(* IEC 61131-3 sources: volt/packages/volt-lsp-iec/test-corpus/bakon-nano/Device/Plc Logic/Application/Library Manager/CAA Callback Extern, 38 files *)

(* ---- CALLBACK.dut ---- *)
TYPE CALLBACK : CB_CALLBACK;
END_TYPE

(* ---- CB_CALLBACK.dut ---- *)
TYPE CB_CALLBACK :
STRUCT
	PPOUFUNC : CAA.PVOID := CAA.gc_pNULL;
	EEVENT : EVENT := EVENT.ALL_EVENTS;
	ECLASS : EVENT_CLASS := EVENT_CLASS.NO_CLASS;
	ESOURCE : EVENT_SOURCE := EVENT_SOURCE.NO_SOURCE;
END_STRUCT
END_TYPE

(* ---- ERROR.dut ---- *)
TYPE ERROR :
(
	NO_ERROR := 0,
	FIRST_ERROR := 20000,
	HANDLE_INVALID := 20001,
	UNKNOWN_EVENT := 20002,
	CALLBACK_NOT_REMOVABLE := 20003,
	WRONG_ARGUMENT := 20004,
	CB_NO_MEMORY := 20005,
	CB_EVENT_EXISTS := 20006,
	CB_CALL_CALLBACKS_FAILED := 20007,
	CB_NO_SYSTEM_EVENT := 20008,
	CB_BUFFER_NOT_AVAILABLE := 20009,
	CB_SYSTEM_EVENT := 20010,
	FIRST_MF := 20050,
	LAST_ERROR := 20099
);
END_TYPE

(* ---- EVENT.dut ---- *)
TYPE EVENT :
(
	ALL_EVENTS := -1,
	NO_EVENT := 0,
	START := 1000,
	STOP,
	BEFORE_RESET,
	AFTER_RESET,
	SHUTDOWN,
	ONLINE_CHANGE,
	BEFORE_DOWNLOAD,
	TASKCODE_NOT_CALLED,
	TIMER,
	DEBUG_LOOP,
	SCHEDULE,
	ERR_WATCHDOG := 4000,
	ERR_HARDWARE_WATCHDOG,
	ERR_FIELDBUS,
	ERR_IOUPDATE,
	ERR_POWERFAIL,
	EXCPT_ILLEGAL_INSTRUCTION := 5000,
	EXCPT_ACCESS_VIOLATION,
	EXCPT_PRIV_INSTRUCTION,
	EXCPT_IN_PAGE_ERROR,
	EXCPT_STACK_OVERFLOW,
	EXCPT_MISALIGNMENT,
	EXCPT_ARRAYBOUNDS,
	EXCPT_DIVIDEBYZERO,
	EXCPT_OVERFLOW,
	EXCPT_NONCONTINUABLE,
	EXCPT_NO_FPU_AVAILABLE := 5500,
	EXCPT_FPU_ERROR,
	EXCPT_FPU_DENORMAL_OPERAND,
	EXCPT_FPU_DIVIDEBYZERO,
	EXCPT_FPU_INVALID_OPERATION,
	EXCPT_FPU_OVERFLOW,
	EXCPT_FPU_STACK_CHECK,
	INTERRUPT_0 := 6000,
	INTERRUPT_1,
	INTERRUPT_2,
	INTERRUPT_3,
	INTERRUPT_4,
	INTERRUPT_5,
	INTERRUPT_6,
	INTERRUPT_7,
	INTERRUPT_8,
	INTERRUPT_9,
	INTERRUPT_10,
	INTERRUPT_11,
	INTERRUPT_12,
	INTERRUPT_13,
	INTERRUPT_14,
	INTERRUPT_15,
	INTERRUPT_255 := 6255,
	AFTER_READING_INPUTS := 7000,
	BEFORE_WRITING_OUTPUTS,
	TIMER_0 := 9900,
	TIMER_1,
	TIMER_2,
	TIMER_3,
	TIMER_4,
	TIMER_5,
	TIMER_6,
	TIMER_7,
	TIMER_8,
	TIMER_9,
	TIMER_10,
	TIMER_11,
	TIMER_12,
	TIMER_13,
	TIMER_14,
	TIMER_15,
	TIMER_99 := 9999
);
END_TYPE

(* ---- EVENT_CLASS.dut ---- *)
TYPE EVENT_CLASS :
(
	ALL_CLASSES := -1,
	NO_CLASS := 16#0,
	ONLINE_EVENTS := 16#1,
	INFOS := 16#2,
	WARNINGS := 16#4,
	RTS_ERRORS := 16#8,
	SYSTEM_EXCEPTIONS := 16#10,
	INTERRUPTS := 16#20,
	IO := 16#40,
	FIELDBUS := 16#80,
	TIMERS := 16#100,
	MANUF_SPEC := 16#200
);
END_TYPE

(* ---- EVENT_SOURCE.dut ---- *)
TYPE EVENT_SOURCE :
(
	ALL_SOURCES := -1,
	NO_SOURCE := 0,
	RUNTIME := 16#1,
	SYSTEM := 16#2,
	IECTASK := 16#4,
	IECPROGRAM := 16#8,
	DRIVER := 16#10
);
END_TYPE

(* ---- GLOBALCONSTANTS.gvl ---- *)
VAR_GLOBAL
	GC_CBNULL : CB_CALLBACK := STRUCT(pPOUFunc := CAA.gc_pNULL, eEvent := EVENT.NO_EVENT, eClass := EVENT_CLASS.NO_CLASS, eSource := EVENT_SOURCE.NO_SOURCE);
END_VAR

(* ---- RSHANDLING.gvl ---- *)
VAR_GLOBAL
	G_CALLBACKCLASS : CallbackClass;
END_VAR

(* ---- VERSIONCONSTANTS.gvl ---- *)
VAR_GLOBAL
	GC_BYVERSION : BYTE := 1;
	GC_VERSION_1 : BYTE := 0;
END_VAR

(* ---- _CALLFUNCTIONBYINDEX.pou ---- *)
FUNCTION _CALLFUNCTIONBYINDEX : __XWORD
VAR_INPUT
	PPOUFUNC : CAA.PVOID;
	DWPARAM1 : __XWORD;
	DWPARAM2 : __XWORD;
	DWPARAM3 : __XWORD;
	PEERROR : POINTER TO ERROR;
END_VAR
END_FUNCTION

(* ---- _DECODECLASS.pou ---- *)
FUNCTION _DECODECLASS : EVENT_CLASS
VAR_INPUT
	DWSPEC : DWORD;
END_VAR
END_FUNCTION

(* ---- _DECODEEVENT.pou ---- *)
FUNCTION _DECODEEVENT : EVENT
VAR_INPUT
	DWSPEC : DWORD;
END_VAR
END_FUNCTION

(* ---- _ENCODESPEC.pou ---- *)
FUNCTION _ENCODESPEC : DWORD
VAR_INPUT
	EEVENT : EVENT;
	ECLASS : EVENT_CLASS;
END_VAR
END_FUNCTION

(* ---- _GETCALLBACK.pou ---- *)
FUNCTION _GETCALLBACK : ERROR
VAR_INPUT
	HHANDLE : CAA.HANDLE;
	PCALLBACK : POINTER TO CB_CALLBACK;
END_VAR
END_FUNCTION

(* ---- _GETHANDLEOFCALLBACK.pou ---- *)
FUNCTION _GETHANDLEOFCALLBACK : CAA.HANDLE
VAR_INPUT
	CTNUMBER : CAA.COUNT;
	PEERROR : POINTER TO ERROR;
END_VAR
END_FUNCTION

(* ---- _GETNUMBERACTIVECALLBACKS.pou ---- *)
FUNCTION _GETNUMBERACTIVECALLBACKS : CAA.COUNT
VAR_INPUT
	PEERROR : POINTER TO ERROR;
END_VAR
END_FUNCTION

(* ---- _ISHANDLEVALID.pou ---- *)
FUNCTION _ISHANDLEVALID : BOOL
VAR_INPUT
	HHANDLE : CAA.HANDLE;
	PEERROR : POINTER TO ERROR;
END_VAR
END_FUNCTION

(* ---- _POSTEVENT.pou ---- *)
FUNCTION _POSTEVENT : ERROR
VAR_INPUT
	EEVENT : EVENT;
	ESOURCE : EVENT_SOURCE;
	DWPARAM : __XWORD;
END_VAR
END_FUNCTION

(* ---- _REGISTERCALLBACK.pou ---- *)
FUNCTION _REGISTERCALLBACK : CAA.HANDLE
VAR_INPUT
	CBNEW : CB_CALLBACK;
	PEERROR : POINTER TO ERROR;
END_VAR
END_FUNCTION

(* ---- _SENDEVENT.pou ---- *)
FUNCTION _SENDEVENT : ERROR
VAR_INPUT
	EEVENT : EVENT;
	ESOURCE : EVENT_SOURCE;
	DWPARAM : __XWORD;
END_VAR
END_FUNCTION

(* ---- _UNREGISTERCALLBACK.pou ---- *)
FUNCTION _UNREGISTERCALLBACK : ERROR
VAR_INPUT
	HHANDLE : CAA.HANDLE;
END_VAR
END_FUNCTION

(* ---- CALLFUNCTIONBYINDEX.pou ---- *)
FUNCTION CALLFUNCTIONBYINDEX : __XWORD
VAR_INPUT
	PPOUFUNC : CAA.PVOID;
	DWPARAM1 : __XWORD;
	DWPARAM2 : __XWORD;
	DWPARAM3 : __XWORD;
	PEERROR : POINTER TO ERROR;
END_VAR
END_FUNCTION

(* ---- DECODECLASS.pou ---- *)
FUNCTION DECODECLASS : EVENT_CLASS
VAR_INPUT
	DWSPEC : DWORD;
END_VAR
END_FUNCTION

(* ---- DECODEEVENT.pou ---- *)
FUNCTION DECODEEVENT : EVENT
VAR_INPUT
	DWSPEC : DWORD;
END_VAR
END_FUNCTION

(* ---- ENCODESPEC.pou ---- *)
FUNCTION ENCODESPEC : DWORD
VAR_INPUT
	EEVENT : EVENT;
	ECLASS : EVENT_CLASS;
END_VAR
END_FUNCTION

(* ---- GETCALLBACK.pou ---- *)
FUNCTION GETCALLBACK : ERROR
VAR_INPUT
	HHANDLE : CAA.HANDLE;
	PCALLBACK : POINTER TO CB_CALLBACK;
END_VAR
END_FUNCTION

(* ---- GETHANDLEOFCALLBACK.pou ---- *)
FUNCTION GETHANDLEOFCALLBACK : CAA.HANDLE
VAR_INPUT
	CTNUMBER : CAA.COUNT;
	PEERROR : POINTER TO ERROR;
END_VAR
END_FUNCTION

(* ---- GETLIBVERSION.pou ---- *)
FUNCTION GETLIBVERSION : VERSION
END_FUNCTION

(* ---- GETLIBVERSIONNUMBER.pou ---- *)
FUNCTION GETLIBVERSIONNUMBER : DWORD
END_FUNCTION

(* ---- GETNUMBERACTIVECALLBACKS.pou ---- *)
FUNCTION GETNUMBERACTIVECALLBACKS : CAA.COUNT
VAR_INPUT
	PEERROR : POINTER TO ERROR;
END_VAR
END_FUNCTION

(* ---- GETSUPPLIERVERSION.pou ---- *)
FUNCTION GETSUPPLIERVERSION : WORD
END_FUNCTION

(* ---- ISHANDLEVALID.pou ---- *)
FUNCTION ISHANDLEVALID : BOOL
VAR_INPUT
	HHANDLE : CAA.HANDLE;
	PEERROR : POINTER TO ERROR;
END_VAR
END_FUNCTION

(* ---- ISLIBRELEASED.pou ---- *)
FUNCTION ISLIBRELEASED : BOOL
END_FUNCTION

(* ---- POSTEVENT.pou ---- *)
FUNCTION POSTEVENT : ERROR
VAR_INPUT
	EEVENT : EVENT;
	ESOURCE : EVENT_SOURCE;
	DWPARAM : __XWORD;
END_VAR
END_FUNCTION

(* ---- REGISTERCALLBACK.pou ---- *)
FUNCTION REGISTERCALLBACK : CAA.HANDLE
VAR_INPUT
	CBNEW : CB_CALLBACK;
	PEERROR : POINTER TO ERROR;
END_VAR
END_FUNCTION

(* ---- SENDEVENT.pou ---- *)
FUNCTION SENDEVENT : ERROR
VAR_INPUT
	EEVENT : EVENT;
	ESOURCE : EVENT_SOURCE;
	DWPARAM : __XWORD;
END_VAR
END_FUNCTION

(* ---- UNREGISTERCALLBACK.pou ---- *)
FUNCTION UNREGISTERCALLBACK : ERROR
VAR_INPUT
	HHANDLE : CAA.HANDLE;
END_VAR
END_FUNCTION

(* ---- CALLBACKCLASS.pou ---- *)
FUNCTION_BLOCK CALLBACKCLASS EXTENDS RSMClass
END_FUNCTION_BLOCK

METHOD CLOSE : RSM.ERROR
VAR_INPUT
	HHANDLE : CAA.HANDLE;
END_VAR
END_METHOD
